FUNCTION_BLOCK tu_pos (* Basic Function Block Type *)
  (* Standard: 61499-2 *)
  (* Version 0.0, 10/23/2026, macie, Schneider Electric, Template *)
  PACKAGE Main;
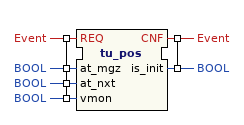
  EVENT_INPUT
    REQ WITH at_mgz, at_nxt, vmon; (* Normal Execution Request *)
  END_EVENT
  EVENT_OUTPUT
    CNF WITH is_init; (* Execution Confirmation *)
  END_EVENT
  VAR_INPUT
    at_mgz : BOOL; (* Input event qualifier *)
    at_nxt : BOOL;
    vmon : BOOL;
  END_VAR
  VAR_OUTPUT
    is_init : BOOL; (* Output event qualifier *)
  END_VAR
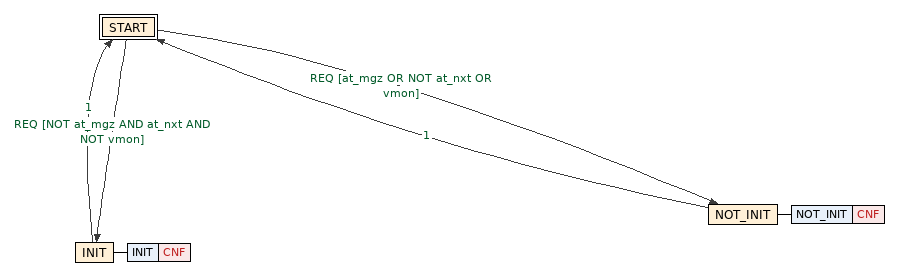
  EC_STATES
    START; (* Initial State *)
    NOT_INIT : NOT_INIT -> CNF; (* Normal execution *)
    INIT : INIT -> CNF;
  END_STATES
  EC_TRANSITIONS
    START TO NOT_INIT := REQ [at_mgz OR NOT at_nxt OR vmon];
    INIT TO START := 1;
    START TO INIT := REQ [NOT at_mgz AND at_nxt AND NOT vmon];
    NOT_INIT TO START := 1;
  END_TRANSITIONS
  ALGORITHM INIT IN ST: (* Initialization algorithm *)
;
is_init := TRUE;
  END_ALGORITHM
  ALGORITHM NOT_INIT IN ST: (* Normally executed algorithm *)
;
is_init := 0;
  END_ALGORITHM
END_FUNCTION_BLOCK
